Fanuc KAREL source: KO00008.KL

PROGRAM KO00008
%NOLOCKGROUP
VAR
  P1: POSITION
  P2: POSITION
  P3: POSITION
  P4: POSITION
  OUT: JOINTPOS
BEGIN
  OUT = FRAME(P1, P2, P3, P4)
END KO00008
